(* CODESYS project listofobject.library
   DefaultNamespace: KOSTAL.TC3.Components.ListOf.Objects
   DocFormat: reStructuredText
   Description: Abstract Class to generate a list of objects.
   Author: Frank Dümpelmann
   Title: KOSTAL.TC3.Components.ListOf.Objects
   Version: 2019.3.1.0
   Company: KOSTAL GmbH & Co.KG
   Placeholder: KOSTAL.TC3.Components.ListOf.Objects

Project tree, tasks and I/O mapping:
  libraries: KOSTAL.TC3.Components.ListOf.Interface, 2019.1.0.0 (KOSTAL GmbH & Co.KG); KOSTAL.TC3.Core.functionResponse, 2019.1.0.0 (KOSTAL GmbH & Co.KG); KOSTAL.TC3.Core.Settings, 2019.0.1.0 (KOSTAL GmbH & Co.KG); KOSTAL.TC3.Core.System, 2019.0.0.0 (KOSTAL GmbH & Co.KG); Tc2_Standard, 3.3.3.0 (Beckhoff Automation GmbH)
  Obsolete/
    V0/
      function block FB_ListOfObject [ST]: AddObject, Clear, New, _DELETE, _deletePayLoad, _New, FB_exit, FB_init
    V1/
      function block FB_Base [ST]: Clear, New, NumberOfObjects, _AddObject, _DELETE, _deletePayLoad, _New, FB_exit, FB_init
      interface I_Base: NumberOfObjects
      interface I_Base_Owner: Clear, New, NumberOfObjects
    data type ST_ListOfObject
  Project Information/
    function F_GetCompany [ST]
    function F_GetTitle [ST]
    function F_GetVersion [ST]
  Version/
    global variables Global_Version
  function block FB_Base_HP [ST]: _removePayload, _verifyMember, _removeMember, _clear, FB_exit, FB_init
  interface I_Base_HP
  interface I_Base_Owner_HP
*)

// Obsolete/ST_ListOfObject
TYPE ST_ListOfObject :
	STRUCT
		pObjects	: POINTER TO PVOID;
		nObjects	: UDINT;
	END_STRUCT
END_TYPE

// Version/Global_Version
{attribute 'TcGenerated'}
{attribute 'no-analysis'}
{attribute 'linkalways'}
// This function has been automatically generated from the project information.
VAR_GLOBAL CONSTANT
	{attribute 'const_non_replaced'}
	stLibVersion_KOSTAL_TC3_Components_ListOf_Objects : ST_LibVersion := (iMajor := 2019, iMinor := 3, iBuild := 1, iRevision := 0, nFlags := 1, sVersion := '2019.3.1.0');
END_VAR

// Obsolete/V0/FB_ListOfObject
{attribute 'obsolete' := 'use instead FB_Base'} 
(*
ListOfObject
============
Abstract Class as Base to create a list of objects with any kind of complex data types.

|-----------------+---------------------------------------------------------------------|
|Parameter        |                                                                     |
|=================+=====================================================================|
|NumberOfElements |defines the number of Objects which shall to create                  | 
|pPVOID           |REFERENCE TO Pointer to a PVOID as Container of all generated Objects| 
|nPVOID           |REFERENCE TO UDINT as Numbers of generated Objects                   | 
|-----------------+---------------------------------------------------------------------|
*)
FUNCTION_BLOCK PUBLIC ABSTRACT FB_ListOfObject

VAR
	_ListOfObject	: ST_ListOfObject;
END_VAR

METHOD PUBLIC AddObject : BOOL;

VAR_INPUT
	ListOfObject			: REFERENCE TO ST_ListOfObject;
END_VAR


VAR
	_u: UDINT;
END_VAR

AddObject:= FALSE;

IF NOT __ISVALIDREF(ListOfObject) THEN RETURN;	END_IF

_ListOfObject.pObjects := 0;
_ListOfObject.nObjects := ListOfObject.nObjects + 1;
_ListOfObject.pObjects:= __NEW(PVOID, _ListOfObject.nObjects);

IF (ListOfObject.pObjects <> 0) AND (ListOfObject.nObjects > 0) THEN 
	FOR _u:= 0 TO ListOfObject.nObjects - 1 DO
		_ListOfObject.pObjects[_u]:= ListOfObject.pObjects[_u];
	END_FOR
END_IF

_ListOfObject.pObjects[_ListOfObject.nObjects - 1]:= _New();

IF (ListOfObject.pObjects <> 0) THEN	__DELETE(ListOfObject.pObjects);	END_IF 

ListOfObject.pObjects:= _ListOfObject.pObjects;
ListOfObject.nObjects:= _ListOfObject.nObjects;

AddObject:= TRUE;
END_METHOD

METHOD PUBLIC Clear
VAR_INPUT
	ListOfObject	: REFERENCE TO ST_ListOfObject;
END_VAR

IF NOT __ISVALIDREF(ListOfObject) THEN RETURN;	END_IF

_ListOfObject.pObjects := ListOfObject.pObjects;
_ListOfObject.nObjects := ListOfObject.nObjects;

_DELETE();

ListOfObject.pObjects:= 0;
ListOfObject.nObjects:= 0;
END_METHOD

METHOD PUBLIC New : BOOL;
VAR_INPUT
	NumberOfElements	: UDINT;
	ListOfObject			: REFERENCE TO ST_ListOfObject;
END_VAR


VAR
	_u: UDINT;
END_VAR

New:= FALSE;

IF NOT __ISVALIDREF(ListOfObject) THEN RETURN;	END_IF

_ListOfObject.pObjects := ListOfObject.pObjects;
_ListOfObject.nObjects := ListOfObject.nObjects;

_DELETE();

IF NumberOfElements = 0 		THEN RETURN;	END_IF

_ListOfObject.nObjects:= NumberOfElements;

_ListOfObject.pObjects:= __NEW(PVOID, _ListOfObject.nObjects);

FOR _u:= 0 TO _ListOfObject.nObjects - 1 DO
	_ListOfObject.pObjects[_u]:= _New();
END_FOR

ListOfObject.pObjects:= _ListOfObject.pObjects;
ListOfObject.nObjects:= _ListOfObject.nObjects;

New:= TRUE;
END_METHOD

METHOD PROTECTED _DELETE

VAR
	_u: UDINT;
END_VAR

IF _ListOfObject.nObjects = 0 THEN 
	IF _ListOfObject.pObjects <> 0 THEN __DELETE(_ListOfObject.pObjects);	END_IF
	RETURN;
END_IF	

IF _ListOfObject.pObjects = 0 THEN _ListOfObject.nObjects:= 0;	RETURN;	END_IF

FOR _u:= 0 TO _ListOfObject.nObjects - 1 DO
	
	_deletePayLoad(_ListOfObject.pObjects[_u]);	
	_ListOfObject.pObjects[_u]:= 0;

END_FOR

IF _ListOfObject.pObjects <> 0 THEN __DELETE(_ListOfObject.pObjects);	END_IF
_ListOfObject.nObjects:= 0;
END_METHOD

//must define in extending FB with real FB-Datatype which is declared with {attribute 'enable_dynamic_creation'}
METHOD PROTECTED ABSTRACT _deletePayLoad
VAR_INPUT
	pPayload	:	PVOID; 
END_VAR
END_METHOD

//must define in extending FB with real FB-Datatype which is declared with {attribute 'enable_dynamic_creation'}
METHOD PROTECTED ABSTRACT _New : PVOID
END_METHOD

METHOD FB_exit : BOOL
VAR_INPUT
	bInCopyCode : BOOL; // if TRUE, the exit method is called for exiting an instance that is copied afterwards (online change).
END_VAR

_DELETE();
END_METHOD

METHOD FB_init : BOOL
VAR_INPUT
	bInitRetains : BOOL; // if TRUE, the retain variables are initialized (warm start / cold start)
	bInCopyCode : BOOL;  // if TRUE, the instance afterwards gets moved into the copy code (online change)
END_VAR

_DELETE();
END_METHOD

END_FUNCTION_BLOCK

// Obsolete/V1/FB_Base
(*
ListOfObject
============
Abstract Class as Base to create a list of objects with any kind of complex data types.
*)
FUNCTION_BLOCK PUBLIC ABSTRACT FB_Base IMPLEMENTS I_Base, I_Base_Owner

VAR
	_ListOfObject	: ST_ListOfObject;
END_VAR

METHOD PUBLIC Clear

_DELETE();

_ListOfObject.pObjects:= 0;
_ListOfObject.nObjects:= 0;
END_METHOD

METHOD PUBLIC New : BOOL;
VAR_INPUT
	NumberOfElements	: UDINT;
END_VAR


VAR
	_u: UDINT;
END_VAR

New:= FALSE;

_DELETE();

IF NumberOfElements = 0 THEN RETURN;	END_IF

_ListOfObject.nObjects:= NumberOfElements;

_ListOfObject.pObjects:= __NEW(PVOID, _ListOfObject.nObjects);

FOR _u:= 0 TO _ListOfObject.nObjects - 1 DO
	_ListOfObject.pObjects[_u]:= _New();
END_FOR

New:= TRUE;
END_METHOD

PROPERTY PUBLIC NumberOfObjects : UDINT
GET

NumberOfObjects:= _ListOfObject.nObjects;
END_GET
END_PROPERTY

//The protected method is used to create a new virtual instance of the class defined in the derived class.
METHOD PROTECTED _AddObject : BOOL;

VAR
	_u: UDINT;
	_copyObj	: ST_ListOfObject;
END_VAR
_AddObject:= FALSE;

_copyObj.pObjects := 0;
_copyObj.nObjects := _ListOfObject.nObjects + 1;
_copyObj.pObjects:= __NEW(PVOID, _copyObj.nObjects);

IF (_ListOfObject.pObjects <> 0) AND (_ListOfObject.nObjects > 0) THEN 
	FOR _u:= 0 TO _ListOfObject.nObjects - 1 DO
		_copyObj.pObjects[_u]:= _ListOfObject.pObjects[_u];
	END_FOR
END_IF

_copyObj.pObjects[_copyObj.nObjects - 1]:= _New();

IF (_ListOfObject.pObjects <> 0) THEN	__DELETE(_ListOfObject.pObjects);	END_IF 

_ListOfObject.pObjects:= _copyObj.pObjects;
_ListOfObject.nObjects:= _copyObj.nObjects;

_AddObject:= TRUE;
END_METHOD

METHOD PROTECTED _DELETE

VAR
	_u: UDINT;
END_VAR

IF _ListOfObject.nObjects = 0 THEN 
	IF _ListOfObject.pObjects <> 0 THEN __DELETE(_ListOfObject.pObjects);	END_IF
	RETURN;
END_IF	

IF _ListOfObject.pObjects = 0 THEN _ListOfObject.nObjects:= 0;	RETURN;	END_IF

FOR _u:= 0 TO _ListOfObject.nObjects - 1 DO
	
	_deletePayLoad(_ListOfObject.pObjects[_u]);	
	_ListOfObject.pObjects[_u]:= 0;

END_FOR

IF _ListOfObject.pObjects <> 0 THEN __DELETE(_ListOfObject.pObjects);	END_IF
_ListOfObject.nObjects:= 0;
END_METHOD

//must define in extending FB with real FB-Datatype which is declared with {attribute 'enable_dynamic_creation'}
METHOD PROTECTED ABSTRACT _deletePayLoad
VAR_INPUT
	pPayload	:	PVOID; 
END_VAR
END_METHOD

//must define in extending FB with real FB-Datatype which is declared with {attribute 'enable_dynamic_creation'}
METHOD PROTECTED ABSTRACT _New : PVOID
END_METHOD

METHOD FB_exit : BOOL
VAR_INPUT
	bInCopyCode : BOOL; // if TRUE, the exit method is called for exiting an instance that is copied afterwards (online change).
END_VAR

_DELETE();
END_METHOD

METHOD FB_init : BOOL
VAR_INPUT
	bInitRetains : BOOL; // if TRUE, the retain variables are initialized (warm start / cold start)
	bInCopyCode : BOOL;  // if TRUE, the instance afterwards gets moved into the copy code (online change)
END_VAR

_DELETE();
END_METHOD

END_FUNCTION_BLOCK

// Obsolete/V1/I_Base
INTERFACE I_Base EXTENDS KOSTAL_TC3_Core_System.I_Interface

PROPERTY PUBLIC NumberOfObjects : UDINT
GET
END_GET
END_PROPERTY

END_INTERFACE

// Obsolete/V1/I_Base_Owner
INTERFACE I_Base_Owner EXTENDS KOSTAL_TC3_Core_System.I_Interface

METHOD PUBLIC Clear
END_METHOD

METHOD PUBLIC New : BOOL;
VAR_INPUT
	NumberOfElements	: UDINT;
END_VAR
END_METHOD

PROPERTY PUBLIC NumberOfObjects : UDINT
GET
END_GET
END_PROPERTY

END_INTERFACE

// Project Information/F_GetCompany
// This function has been automatically generated from the project information.
{attribute 'signature_flag' := '1073741824'}
{attribute 'TcGenerated'}
{attribute 'no-analysis'}
FUNCTION F_GetCompany : WSTRING
VAR_INPUT
	
END_VAR

F_GetCompany := "KOSTAL GmbH & Co.KG";

END_FUNCTION

// Project Information/F_GetTitle
// This function has been automatically generated from the project information.
{attribute 'signature_flag' := '1073741824'}
{attribute 'TcGenerated'}
{attribute 'no-analysis'}
FUNCTION F_GetTitle : WSTRING
VAR_INPUT
	
END_VAR

F_GetTitle := "KOSTAL.TC3.Components.ListOf.Objects";

END_FUNCTION

// Project Information/F_GetVersion
// This function has been automatically generated from the project information.
{attribute 'signature_flag' := '1073741824'}
{attribute 'TcGenerated'}
{attribute 'no-analysis'}
FUNCTION F_GetVersion : ST_LibVersion
VAR_INPUT
	
END_VAR

F_GetVersion.iMajor := 2019;
F_GetVersion.iMinor := 3;
F_GetVersion.iBuild := 1;
F_GetVersion.iRevision := 0;
F_GetVersion.sVersion := '2019.3.1.0';
F_GetVersion.nFlags := 1;

END_FUNCTION

// FB_Base_HP
(*

| ==================================================================================
| List of Items of objects with base Interface {KOSTAL_TC3_Core_System.I_Interface} 
| ==================================================================================

..code::

	//In addition to the interface, each item contains the pointer to the previous item 
	//as well as the pointer to the next item in the list.

	TYPE ST_List :
		STRUCT
				pNext			: P_List;
				iMember		: KOSTAL_TC3_Core_System.I_Interface;	
				pPrevious : P_List;
		END_STRUCT
	END_TYPE

============= ======================================= ======================
| The List is defined by (p)Begin and (p)End and also the count of Members 
----------------------------------------------------------------------------
============= ======================================= ======================
 **_pBegin**  >>>>>>>>>>>>>>>>>>>>>>>>>>>>>>>>>>>>>>  **_pEnd**                     
 **Item-1**	    Item-2   Item-3   Item-4  Item-5      **Item-n**                   
============= ======================================= ======================



| =========================================================================
| The Member is an object which implements the base Interface as payload. 
| -------------------------------------------------------------------------
| Previous Item ---<<<Pointer-Previous-[Item]-Pointer-Next>>>---NextItem---
| =========================================================================

*)
FUNCTION_BLOCK ABSTRACT FB_Base_HP EXTENDS KOSTAL_TC3_Components_ListOf_Interface.FB_Base IMPLEMENTS I_Base_HP, I_Base_Owner_HP

(*
	Integrate the type-specific procedures here to clean up the member and remove it from memory. 
	only if verifing is passed [_verifyMember:= TRUE] the called metode should proceed 
*)
METHOD PROTECTED _removePayload : BOOL
VAR_INPUT
	Member	: KOSTAL_TC3_Core_System.I_Interface;
	Result	: REFERENCE TO KOSTAL_TC3_Core_functionResponse.FB_functionResponse;
END_VAR

_removePayload:= TRUE;
END_METHOD

(*
	integrate here the veryfing of your interface type 
	only if verifing is passed [_verifyMember:= TRUE] the called metode will proceeded 
*)
METHOD PROTECTED _verifyMember : BOOL

VAR_INPUT
	Member	: KOSTAL_TC3_Core_System.I_Interface;
	Result	: REFERENCE TO KOSTAL_TC3_Core_functionResponse.FB_functionResponse;
END_VAR

VAR
	_obj	: KOSTAL_TC3_Core_System.I_Interface;
	_bResult: BOOL;
END_VAR

IF Member = 0 THEN _setResultFail(Result, 'Parameter Member is empty');	RETURN;	END_IF

_bResult:= __QUERYINTERFACE(Member, _obj);

IF NOT _bResult OR (_obj = 0) THEN
	IF __ISVALIDREF(Result) THEN Result.success:= FALSE; Result.status:= 'no valid interface found';	END_IF	
	RETURN;
END_IF

_verifyMember:= TRUE;
END_METHOD

(*
	remove given {Member} from List including the customer payload {_removePayload()]
*)
METHOD PROTECTED _removeMember : BOOL
VAR_INPUT
	Member	: KOSTAL_TC3_Core_System.I_Interface;
	Result	: REFERENCE TO KOSTAL_TC3_Core_functionResponse.FB_functionResponse;
END_VAR

VAR
	_Item		: P_List;
	_bFound: BOOL;
END_VAR
IF NOT _verifyMember(Member, Result)	THEN	RETURN;	END_IF

_bFound:= _findItem(Member, _Item, Result);

IF NOT _bFound THEN RETURN;	END_IF

_removePayload(Member, Result);

_removeMember:= _removeItem(_Item, Result);
END_METHOD

(*
	Delete the complete content of the list including the customer payload {_removePayload()}
*)
METHOD PROTECTED _clear

WHILE THIS^._pBegin <> 0 DO
	_removePayload(THIS^._pBegin^.iMember, 0);
  THIS^._removeMember(THIS^._pBegin^.iMember, 0);  
END_WHILE
END_METHOD

METHOD FB_exit : BOOL
VAR_INPUT
	bInCopyCode : BOOL; // if TRUE, the exit method is called for exiting an instance that is copied afterwards (online change).
END_VAR

_clear();
END_METHOD

METHOD FB_init : BOOL
VAR_INPUT
	bInitRetains : BOOL; // if TRUE, the retain variables are initialized (warm start / cold start)
	bInCopyCode : BOOL;  // if TRUE, the instance afterwards gets moved into the copy code (online change)
END_VAR

_clear();
END_METHOD

END_FUNCTION_BLOCK

// I_Base_HP
INTERFACE I_Base_HP EXTENDS KOSTAL_TC3_Components_ListOf_Interface.I_Base

END_INTERFACE

// I_Base_Owner_HP
INTERFACE I_Base_Owner_HP EXTENDS KOSTAL_TC3_Components_ListOf_Interface.I_Base_Owner

END_INTERFACE
